Fanuc KAREL source: kt00146.KL

-- PROVISIONAL review KL for V770-1; original PC SHA256 ef17c019e0be768541f0c9f47866f4a317f7c31ce6530fa138f489701c31b576
-- Incomplete behavior may be omitted. Consult companion uncertainty JSON. Do not deploy.
PROGRAM KT00146
%NOLOCKGROUP
VAR
  I2 : INTEGER
  OUT : REAL
-- UNRESOLVED_DECL Y1 type=002018
BEGIN
  -- UNRESOLVED_PC offsets 5-19; opcodes 2E,22,9D,33,B2
  -- UNRESOLVED_PC offsets 24-35; opcodes 2E,23
  -- UNRESOLVED_PC offsets 40-63; opcodes 22,9D,33,B1,21,55,64,23
  -- UNRESOLVED_PC offsets 68-72; opcodes 7F
END KT00146
